(* IEC 61131-3 sources: guidance-for-physical-ai-production-designer-on-aws/source/plan2cell/crates/bt2plc/tests/golden/cell_2robot/codesys/head/GVL, 2 files *)

(* ---- GVL_Cell.st ---- *)
(*
 * GVL_Cell - generated by bt2plc 0.1.0 - DO NOT EDIT
 * Plan   : bt_1791274820_cell_2robot (cell cell_2robot)
 * Grants : planned ticket order
 *)
{attribute 'qualified_only'}
VAR_GLOBAL CONSTANT
    (* ========================================================================
       DIMENSIONS (array bounds are literals; *_DIM >= 1)
       ======================================================================== *)
    N_ROBOTS                : INT := 1;
    N_ZONES                 : INT := 0;
    N_OPS                   : INT := 2;
    N_PREDS                 : INT := 0;

    (* ========================================================================
       PROTOCOL / TIMING
       ======================================================================== *)
    PLAN_ID                 : WORD := WORD#16#A312;             (* fold of the plan fingerprint *)
    PROD_FOLGE              : WORD := WORD#11;                  (* default production Folge *)
    HOME_FOLGE              : WORD := WORD#125;                 (* blind homing *)
    JOB_NUMBER_BYTE         : BOOL := FALSE;                    (* FALSE: WORD LE bytes 2-3, TRUE: byte 2 *)
    PROFILE_VW              : BOOL := FALSE;                    (* TRUE: VW KS24 signal map and Folge handshake instead of the simulator telegram *)
    GRANT_POLICY            : E_GrantPolicy := E_GrantPolicy.GP_PLANNED;
    HOME_SEQUENTIAL         : BOOL := TRUE;
    AUTO_RUN                : BOOL := TRUE;                     (* start the next cycle automatically *)
    STEP_BYTE               : INT := 4;                         (* robot -> PLC, WORD LE op index *)
    REQ_BYTE                : INT := 28;                        (* robot -> PLC, DWORD LE zone requests *)
    GRANT_BYTE              : INT := 12;                        (* PLC -> robot, DWORD LE zone grants *)
    PLAN_ID_BYTE            : INT := 4;                         (* PLC -> robot, WORD LE plan id *)
    PERMIT_MASK             : DWORD := DWORD#16#80000000;       (* bit 31: permit predecessors *)
    T_RESET_PULSE           : TIME := T#1S;
    T_START_PULSE           : TIME := T#500MS;
    T_STOP_PULSE            : TIME := T#1S;
    T_HANDSHAKE             : TIME := T#5S;
    T_BRINGUP_LIMIT         : TIME := T#1M;                     (* safety enable: PROFINET connection set-up *)
    T_MISMATCH_DEBOUNCE     : TIME := T#200MS;
    T_STOP_DEBOUNCE         : TIME := T#200MS;                  (* job running: ProgRunning and ProgFinished low this long = robot stopped *)
    T_CYCLE_PAUSE           : TIME := T#2S;
    T_START_LIMIT           : TIME := T#15S;
    T_ABORT_LIMIT           : TIME := T#10S;
    T_HOME_LIMIT            : TIME := T#15S500MS;

    (* ========================================================================
       VW KS24 SIGNAL INDICES (used when PROFILE_VW; $IN/$OUT index, 1-based)
       ======================================================================== *)
    VW_READY_OUT            : INT := 9;                         (* O_R_Bereit *)
    VW_RK100_OUT            : INT := 10;                        (* O_R_RK100 safety circuit *)
    VW_AUTO_OUT             : INT := 12;                        (* O_R_Auto *)
    VW_ESTOP_OUT            : INT := 13;                        (* O_R_Notaus *)
    VW_END_OUT              : INT := 14;                        (* O_R_F_ENDE / LPKT *)
    VW_PF0_OUT              : INT := 15;                        (* O_R_PFO home position *)
    VW_STEP_OUT             : INT := 97;                        (* P_PktNr_SPS op index (16 bits) *)
    VW_REL_OUT              : INT := 41;                        (* interlock releases A41-56 *)
    VW_REQ_OUT              : INT := 81;                        (* interlock requests A81-96 *)
    VW_ERR_OUT              : INT := 225;                       (* VW_FEH_BIN_A error code (8 bits) *)
    VW_DRIVES_IN            : INT := 10;                        (* I_R_Ant_Ein *)
    VW_SRB_IN               : INT := 9;                         (* I_R_SRB Folge start *)
    VW_RESET_IN             : INT := 26;                        (* I_R_Quit_St acknowledge *)
    anInterlock             : ARRAY[1..1] OF INT := [0];        (* robot r, zone z -> VW interlock 1..16 (0 = not a member): index (r-1)*1+z *)

    (* ========================================================================
       ROBOTS (index = BT order)
       ======================================================================== *)
    asRobotTag              : ARRAY[1..1] OF STRING(16) := ['R1'];
    asRobotNs               : ARRAY[1..1] OF STRING(32) := ['robot1'];
    abRobotActive           : ARRAY[1..1] OF BOOL := [TRUE];
    abSafetyBypass          : ARRAY[1..1] OF BOOL := [FALSE];   (* SIMULATION ONLY: PROFIsafe slot-1 bits not required ([[robot]] safety_bypass) *)
    awRobotProdFolge        : ARRAY[1..1] OF WORD := [WORD#11];
    anRobotFirstOp          : ARRAY[1..1] OF INT := [1];        (* op k of robot r: aOps[anRobotFirstOp[r] + k - 1] *)
    anRobotOpCount          : ARRAY[1..1] OF INT := [2];

    (* ========================================================================
       ZONES - tickets of zone z: aTickets[anZoneFirst[z] .. anZoneFirst[z] + anZoneCount[z] - 1]
       ======================================================================== *)
    asZoneName              : ARRAY[1..1] OF STRING(8) := [''];
    anZoneFirst             : ARRAY[1..1] OF INT := [0];
    anZoneCount             : ARRAY[1..1] OF INT := [0];
    aTickets                : ARRAY[1..1] OF ST_Ticket := [
        (nRobot := 0, nOp := 0)    (* no zones *)
    ];

    (* ========================================================================
       OPS - op k of robot r: aOps[anRobotFirstOp[r] + k - 1]
       ======================================================================== *)
    (* tLimit = 1.5 x tExpected + 5 s ; tZoneDeadline = 1.5 x ASAP grant + (5 + 0.2) s x depth + 10 s *)
    aOps                    : ARRAY[1..2] OF ST_OpInfo := [
        (nRobot := 1, nOp := 1, dwZoneMask := DWORD#16#00000000, nPredFirst := 0, nPredCount := 0, tExpected := T#3S729MS, tLimit := T#10S594MS, tZoneDeadline := T#10S, sName := 'STAGE_R1'),    (* R1 #1 STAGE_R1 *)
        (nRobot := 1, nOp := 2, dwZoneMask := DWORD#16#00000000, nPredFirst := 0, nPredCount := 0, tExpected := T#2S419MS, tLimit := T#8S629MS, tZoneDeadline := T#20S794MS, sName := 'HOME')    (* R1 #2 HOME *)
    ];

    (* ========================================================================
       PERMIT PREDECESSORS - op preds: aPreds[nPredFirst .. nPredFirst + nPredCount - 1]
       ======================================================================== *)
    aPreds                  : ARRAY[1..1] OF ST_Ticket := [
        (nRobot := 0, nOp := 0)    (* no permit predecessors *)
    ];
END_VAR

(* ---- GVL_IO.st ---- *)
(*
 * GVL_IO - Head PLC I/O, one block per robot
 * Generated by bt2plc 0.1.0 for cell cell_2robot (plan bt_1791274820_cell_2robot)
 *
 * This is the PROFINET Controller (master) side.
 * From the controller's perspective:
 *   "Inputs"  = data received FROM the robot device (robot status)
 *   "Outputs" = data sent TO the robot device (PLC commands)
 *
 * Map in the I/O Mapping tab of each KUKA device under the PN-Controller:
 *   SafeIO_FDIO64_<tag> inputs  -> bySafeIn0_<tag>..bySafeIn7_<tag>
 *   SafeIO_FDIO64_<tag> outputs -> bySafeOut0_<tag>..bySafeOut7_<tag>
 *   VASS_DIO256_<tag> inputs    -> aVassInputData_<tag>
 *   VASS_DIO256_<tag> outputs   -> aVassOutputData_<tag>
 *
 * Only PLC_PRG accesses this GVL: whole arrays and single bytes are copied
 * into / out of FB_Cell (never write single elements of these arrays).
 *)

{attribute 'qualified_only'}
VAR_GLOBAL

    (* ========================================================================
       R1 - robot1 - kuka_robi1 (kuka-robi1, 192.168.100.11)
       ======================================================================== *)

    (* SLOT 1 - PROFIsafe FDIO64: safe status FROM robot (8 bytes) *)
    bySafeIn0_R1            : BYTE;     (* Byte 0: Drives OK, Stopped, Reduced speed... *)
    bySafeIn1_R1            : BYTE;     (* Byte 1: Gates, E-Stop, Enabling... *)
    bySafeIn2_R1            : BYTE;     (* Byte 2: STO, SS1, SS2, SOS, SLS... *)
    bySafeIn3_R1            : BYTE;
    bySafeIn4_R1            : BYTE;
    bySafeIn5_R1            : BYTE;
    bySafeIn6_R1            : BYTE;
    bySafeIn7_R1            : BYTE;

    (* SLOT 1 - PROFIsafe FDIO64: safe commands TO robot (8 bytes) *)
    bySafeOut0_R1           : BYTE;     (* Byte 0: Drive enable, E-Stop, SS1, SS2, SLS... *)
    bySafeOut1_R1           : BYTE;     (* Byte 1: Zone enables *)
    bySafeOut2_R1           : BYTE;
    bySafeOut3_R1           : BYTE;
    bySafeOut4_R1           : BYTE;
    bySafeOut5_R1           : BYTE;
    bySafeOut6_R1           : BYTE;
    bySafeOut7_R1           : BYTE;

    (* SLOT 2 - DIO256 VASS telegram (32 bytes each direction) *)
    aVassInputData_R1       : ARRAY[0..31] OF BYTE;         (* VASS status FROM robot *)
    aVassOutputData_R1      : ARRAY[0..31] OF BYTE;         (* VASS commands TO robot *)

END_VAR
